TYPE ST_Cia402Drive :
STRUCT
    // Drive to PLC (TxPDO): copy in before each call. All three needed.
    nStatusword       : WORD;   // 0x6041
    nModesDisplay     : SINT;   // 0x6061
    nPositionActual   : DINT;   // 0x6064
    // PLC to drive (RxPDO): copy out after each call.
    nControlword      : WORD;   // 0x6040, written by the FB only
    nModesOfOperation : SINT;   // 0x6060, written by the FB only
    nTargetPosition   : DINT;   // 0x607A
    nTargetVelocity   : DINT;   // 0x60FF
    nTargetTorque     : INT;    // 0x6071
    // Caller to FB: controlword bits 4-6, 8, 9, sent only while bValid.
    nModeBits         : WORD;
END_STRUCT
END_TYPE

(* stored: Version 1.1.0.1, ProductVersion 3.1.4024.0
   DUT ST_Cia402Drive: Id {1ef61cea-b0b3-4865-ae01-9923f3d96540} *)
